Fanuc KAREL source: KB00055.KL

PROGRAM KB00055
%NOLOCKGROUP
VAR
  P1: INTEGER
  P2: INTEGER
  P3: STRING[80]
  P4: INTEGER
BEGIN
  P1 = 1
  P2 = 1
  P3 = 'A'
  P4 = 1
  DAQ_START(P1, P2, P3, P4)
END KB00055
